Fanuc KAREL source: KT00924.KL

PROGRAM KT00924
%NOLOCKGROUP
VAR
  I1: INTEGER
  I2: INTEGER
  OUT: STRING[80]
BEGIN
  I1 = 2
  I2 = 3
  I1 = 2
  I2 = 3
  OUT = SUB_STR(I1, 1, 1)
END KT00924
